Universal Robots URScript: horizontal_swab_path 7.script

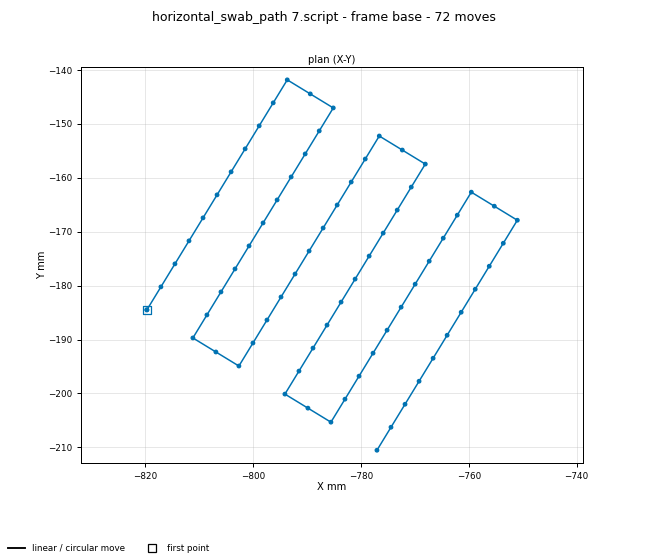
[picture p0: tool path of horizontal_swab_path 7.script in frame base, 72 of 72 moves have a stored position in this frame; points joined in program order, loops and branches not executed]
def horizontal_swab_path():

  # Move to first swab point perpendicular
  movel(p[-0.81971797, -0.18449305, 0.03056454, 2.72713527, 1.53061624, -0.02224013], a=0.2000, v=0.0300, r=0.0000)

  # Incline tool while keeping TCP XYZ fixed
  movel(p[-0.81971797, -0.18449305, 0.03056454, -2.11716639, -1.17714539, 0.50774966], a=0.1000, v=0.0150, r=0.0000)
  # Horizontal waypoint 1
  movel(p[-0.81711371, -0.18022591, 0.03046777, -2.11716639, -1.17714539, 0.50774966], a=0.1500, v=0.0200, r=0.0100)
  # Horizontal waypoint 2
  movel(p[-0.81450945, -0.17595878, 0.03037099, -2.11716639, -1.17714539, 0.50774966], a=0.1500, v=0.0200, r=0.0100)
  # Horizontal waypoint 3
  movel(p[-0.81190518, -0.17169164, 0.03027422, -2.11716639, -1.17714539, 0.50774966], a=0.1500, v=0.0200, r=0.0100)
  # Horizontal waypoint 4
  movel(p[-0.80930092, -0.16742450, 0.03017745, -2.11716639, -1.17714539, 0.50774966], a=0.1500, v=0.0200, r=0.0100)
  # Horizontal waypoint 5
  movel(p[-0.80669666, -0.16315737, 0.03008068, -2.11716639, -1.17714539, 0.50774966], a=0.1500, v=0.0200, r=0.0100)
  # Horizontal waypoint 6
  movel(p[-0.80409240, -0.15889023, 0.02998390, -2.11716639, -1.17714539, 0.50774966], a=0.1500, v=0.0200, r=0.0100)
  # Horizontal waypoint 7
  movel(p[-0.80148814, -0.15462309, 0.02988713, -2.11716639, -1.17714539, 0.50774966], a=0.1500, v=0.0200, r=0.0100)
  # Horizontal waypoint 8
  movel(p[-0.79888387, -0.15035596, 0.02979036, -2.11716639, -1.17714539, 0.50774966], a=0.1500, v=0.0200, r=0.0100)
  # Horizontal waypoint 9
  movel(p[-0.79627961, -0.14608882, 0.02969359, -2.11716639, -1.17714539, 0.50774966], a=0.1500, v=0.0200, r=0.0100)
  # Horizontal waypoint 10
  movel(p[-0.79367535, -0.14182168, 0.02959681, -2.11716639, -1.17714539, 0.50774966], a=0.1500, v=0.0200, r=0.0100)
  # Horizontal waypoint 11
  movel(p[-0.78940720, -0.14442595, 0.02962395, -2.11716639, -1.17714539, 0.50774966], a=0.1500, v=0.0200, r=0.0100)
  # Horizontal waypoint 12
  movel(p[-0.78513906, -0.14703021, 0.02965108, -2.11716639, -1.17714539, 0.50774966], a=0.1500, v=0.0200, r=0.0100)
  # Horizontal waypoint 13
  movel(p[-0.78774332, -0.15129735, 0.02974786, -2.11716639, -1.17714539, 0.50774966], a=0.1500, v=0.0200, r=0.0100)
  # Horizontal waypoint 14
  movel(p[-0.79034758, -0.15556448, 0.02984463, -2.11716639, -1.17714539, 0.50774966], a=0.1500, v=0.0200, r=0.0100)
  # Horizontal waypoint 15
  movel(p[-0.79295184, -0.15983162, 0.02994140, -2.11716639, -1.17714539, 0.50774966], a=0.1500, v=0.0200, r=0.0100)
  # Horizontal waypoint 16
  movel(p[-0.79555610, -0.16409876, 0.03003817, -2.11716639, -1.17714539, 0.50774966], a=0.1500, v=0.0200, r=0.0100)
  # Horizontal waypoint 17
  movel(p[-0.79816037, -0.16836589, 0.03013494, -2.11716639, -1.17714539, 0.50774966], a=0.1500, v=0.0200, r=0.0100)
  # Horizontal waypoint 18
  movel(p[-0.80076463, -0.17263303, 0.03023172, -2.11716639, -1.17714539, 0.50774966], a=0.1500, v=0.0200, r=0.0100)
  # Horizontal waypoint 19
  movel(p[-0.80336889, -0.17690016, 0.03032849, -2.11716639, -1.17714539, 0.50774966], a=0.1500, v=0.0200, r=0.0100)
  # Horizontal waypoint 20
  movel(p[-0.80597315, -0.18116730, 0.03042526, -2.11716639, -1.17714539, 0.50774966], a=0.1500, v=0.0200, r=0.0100)
  # Horizontal waypoint 21
  movel(p[-0.80857742, -0.18543444, 0.03052203, -2.11716639, -1.17714539, 0.50774966], a=0.1500, v=0.0200, r=0.0100)
  # Horizontal waypoint 22
  movel(p[-0.81118168, -0.18970158, 0.03061881, -2.11716639, -1.17714539, 0.50774966], a=0.1500, v=0.0200, r=0.0100)
  # Horizontal waypoint 23
  movel(p[-0.80691353, -0.19230584, 0.03064594, -2.11716639, -1.17714539, 0.50774966], a=0.1500, v=0.0200, r=0.0100)
  # Horizontal waypoint 24
  movel(p[-0.80264539, -0.19491010, 0.03067308, -2.11716639, -1.17714539, 0.50774966], a=0.1500, v=0.0200, r=0.0100)
  # Horizontal waypoint 25
  movel(p[-0.80004112, -0.19064296, 0.03057630, -2.11716639, -1.17714539, 0.50774966], a=0.1500, v=0.0200, r=0.0100)
  # Horizontal waypoint 26
  movel(p[-0.79743686, -0.18637583, 0.03047953, -2.11716639, -1.17714539, 0.50774966], a=0.1500, v=0.0200, r=0.0100)
  # Horizontal waypoint 27
  movel(p[-0.79483260, -0.18210869, 0.03038276, -2.11716639, -1.17714539, 0.50774966], a=0.1500, v=0.0200, r=0.0100)
  # Horizontal waypoint 28
  movel(p[-0.79222834, -0.17784156, 0.03028599, -2.11716639, -1.17714539, 0.50774966], a=0.1500, v=0.0200, r=0.0100)
  # Horizontal waypoint 29
  movel(p[-0.78962407, -0.17357442, 0.03018921, -2.11716639, -1.17714539, 0.50774966], a=0.1500, v=0.0200, r=0.0100)
  # Horizontal waypoint 30
  movel(p[-0.78701981, -0.16930728, 0.03009244, -2.11716639, -1.17714539, 0.50774966], a=0.1500, v=0.0200, r=0.0100)
  # Horizontal waypoint 31
  movel(p[-0.78441555, -0.16504015, 0.02999567, -2.11716639, -1.17714539, 0.50774966], a=0.1500, v=0.0200, r=0.0100)
  # Horizontal waypoint 32
  movel(p[-0.78181129, -0.16077301, 0.02989890, -2.11716639, -1.17714539, 0.50774966], a=0.1500, v=0.0200, r=0.0100)
  # Horizontal waypoint 33
  movel(p[-0.77920703, -0.15650587, 0.02980212, -2.11716639, -1.17714539, 0.50774966], a=0.1500, v=0.0200, r=0.0100)
  # Horizontal waypoint 34
  movel(p[-0.77660276, -0.15223874, 0.02970535, -2.11716639, -1.17714539, 0.50774966], a=0.1500, v=0.0200, r=0.0100)
  # Horizontal waypoint 35
  movel(p[-0.77233462, -0.15484300, 0.02973249, -2.11716639, -1.17714539, 0.50774966], a=0.1500, v=0.0200, r=0.0100)
  # Horizontal waypoint 36
  movel(p[-0.76806647, -0.15744726, 0.02975962, -2.11716639, -1.17714539, 0.50774966], a=0.1500, v=0.0200, r=0.0100)
  # Horizontal waypoint 37
  movel(p[-0.77067073, -0.16171440, 0.02985639, -2.11716639, -1.17714539, 0.50774966], a=0.1500, v=0.0200, r=0.0100)
  # Horizontal waypoint 38
  movel(p[-0.77327499, -0.16598154, 0.02995317, -2.11716639, -1.17714539, 0.50774966], a=0.1500, v=0.0200, r=0.0100)
  # Horizontal waypoint 39
  movel(p[-0.77587926, -0.17024867, 0.03004994, -2.11716639, -1.17714539, 0.50774966], a=0.1500, v=0.0200, r=0.0100)
  # Horizontal waypoint 40
  movel(p[-0.77848352, -0.17451581, 0.03014671, -2.11716639, -1.17714539, 0.50774966], a=0.1500, v=0.0200, r=0.0100)
  # Horizontal waypoint 41
  movel(p[-0.78108778, -0.17878295, 0.03024348, -2.11716639, -1.17714539, 0.50774966], a=0.1500, v=0.0200, r=0.0100)
  # Horizontal waypoint 42
  movel(p[-0.78369204, -0.18305008, 0.03034026, -2.11716639, -1.17714539, 0.50774966], a=0.1500, v=0.0200, r=0.0100)
  # Horizontal waypoint 43
  movel(p[-0.78629631, -0.18731722, 0.03043703, -2.11716639, -1.17714539, 0.50774966], a=0.1500, v=0.0200, r=0.0100)
  # Horizontal waypoint 44
  movel(p[-0.78890057, -0.19158436, 0.03053380, -2.11716639, -1.17714539, 0.50774966], a=0.1500, v=0.0200, r=0.0100)
  # Horizontal waypoint 45
  movel(p[-0.79150483, -0.19585149, 0.03063057, -2.11716639, -1.17714539, 0.50774966], a=0.1500, v=0.0200, r=0.0100)
  # Horizontal waypoint 46
  movel(p[-0.79410909, -0.20011863, 0.03072735, -2.11716639, -1.17714539, 0.50774966], a=0.1500, v=0.0200, r=0.0100)
  # Horizontal waypoint 47
  movel(p[-0.78984095, -0.20272289, 0.03075448, -2.11716639, -1.17714539, 0.50774966], a=0.1500, v=0.0200, r=0.0100)
  # Horizontal waypoint 48
  movel(p[-0.78557280, -0.20532716, 0.03078161, -2.11716639, -1.17714539, 0.50774966], a=0.1500, v=0.0200, r=0.0100)
  # Horizontal waypoint 49
  movel(p[-0.78296854, -0.20106002, 0.03068484, -2.11716639, -1.17714539, 0.50774966], a=0.1500, v=0.0200, r=0.0100)
  # Horizontal waypoint 50
  movel(p[-0.78036428, -0.19679288, 0.03058807, -2.11716639, -1.17714539, 0.50774966], a=0.1500, v=0.0200, r=0.0100)
  # Horizontal waypoint 51
  movel(p[-0.77776001, -0.19252575, 0.03049130, -2.11716639, -1.17714539, 0.50774966], a=0.1500, v=0.0200, r=0.0100)
  # Horizontal waypoint 52
  movel(p[-0.77515575, -0.18825861, 0.03039452, -2.11716639, -1.17714539, 0.50774966], a=0.1500, v=0.0200, r=0.0100)
  # Horizontal waypoint 53
  movel(p[-0.77255149, -0.18399147, 0.03029775, -2.11716639, -1.17714539, 0.50774966], a=0.1500, v=0.0200, r=0.0100)
  # Horizontal waypoint 54
  movel(p[-0.76994723, -0.17972434, 0.03020098, -2.11716639, -1.17714539, 0.50774966], a=0.1500, v=0.0200, r=0.0100)
  # Horizontal waypoint 55
  movel(p[-0.76734296, -0.17545720, 0.03010421, -2.11716639, -1.17714539, 0.50774966], a=0.1500, v=0.0200, r=0.0100)
  # Horizontal waypoint 56
  movel(p[-0.76473870, -0.17119006, 0.03000744, -2.11716639, -1.17714539, 0.50774966], a=0.1500, v=0.0200, r=0.0100)
  # Horizontal waypoint 57
  movel(p[-0.76213444, -0.16692293, 0.02991066, -2.11716639, -1.17714539, 0.50774966], a=0.1500, v=0.0200, r=0.0100)
  # Horizontal waypoint 58
  movel(p[-0.75953018, -0.16265579, 0.02981389, -2.11716639, -1.17714539, 0.50774966], a=0.1500, v=0.0200, r=0.0100)
  # Horizontal waypoint 59
  movel(p[-0.75526203, -0.16526005, 0.02984103, -2.11716639, -1.17714539, 0.50774966], a=0.1500, v=0.0200, r=0.0100)
  # Horizontal waypoint 60
  movel(p[-0.75099388, -0.16786432, 0.02986816, -2.11716639, -1.17714539, 0.50774966], a=0.1500, v=0.0200, r=0.0100)
  # Horizontal waypoint 61
  movel(p[-0.75359814, -0.17213145, 0.02996493, -2.11716639, -1.17714539, 0.50774966], a=0.1500, v=0.0200, r=0.0100)
  # Horizontal waypoint 62
  movel(p[-0.75620241, -0.17639859, 0.03006171, -2.11716639, -1.17714539, 0.50774966], a=0.1500, v=0.0200, r=0.0100)
  # Horizontal waypoint 63
  movel(p[-0.75880667, -0.18066573, 0.03015848, -2.11716639, -1.17714539, 0.50774966], a=0.1500, v=0.0200, r=0.0100)
  # Horizontal waypoint 64
  movel(p[-0.76141093, -0.18493286, 0.03025525, -2.11716639, -1.17714539, 0.50774966], a=0.1500, v=0.0200, r=0.0100)
  # Horizontal waypoint 65
  movel(p[-0.76401520, -0.18920000, 0.03035202, -2.11716639, -1.17714539, 0.50774966], a=0.1500, v=0.0200, r=0.0100)
  # Horizontal waypoint 66
  movel(p[-0.76661946, -0.19346714, 0.03044880, -2.11716639, -1.17714539, 0.50774966], a=0.1500, v=0.0200, r=0.0100)
  # Horizontal waypoint 67
  movel(p[-0.76922372, -0.19773427, 0.03054557, -2.11716639, -1.17714539, 0.50774966], a=0.1500, v=0.0200, r=0.0100)
  # Horizontal waypoint 68
  movel(p[-0.77182798, -0.20200141, 0.03064234, -2.11716639, -1.17714539, 0.50774966], a=0.1500, v=0.0200, r=0.0100)
  # Horizontal waypoint 69
  movel(p[-0.77443224, -0.20626855, 0.03073911, -2.11716639, -1.17714539, 0.50774966], a=0.1500, v=0.0200, r=0.0100)
  # Horizontal waypoint 70
  movel(p[-0.77703651, -0.21053568, 0.03083589, -2.11716639, -1.17714539, 0.50774966], a=0.1500, v=0.0200, r=0.0100)

end
